TYPE "ST_CommandInfo"
VERSION : 0.1
   STRUCT
      "Value" : DInt;
      "Label" : String[120];
      "Style" : DInt;
   END_STRUCT;
END_TYPE
